Fanuc KAREL source: kt00881.KL

-- PROVISIONAL review KL for V770-1; original PC SHA256 7bfcebda0242e58e16e4d91c53400874c8d9c3006e6fad8e13b8db4fe4a92cd5
-- Incomplete behavior may be omitted. Consult companion uncertainty JSON. Do not deploy.
PROGRAM KT00881
%NOLOCKGROUP
VAR
  I1 : INTEGER
  I2 : INTEGER
  OUT : REAL
BEGIN
  -- UNRESOLVED_PC offsets 5-16; opcodes 2E,23
  -- UNRESOLVED_PC offsets 21-32; opcodes 2E,23
  -- UNRESOLVED_PC offsets 37-48; opcodes 2E,23
  -- UNRESOLVED_PC offsets 53-64; opcodes 2E,23
  -- UNRESOLVED_PC offsets 69-94; opcodes 27,27,21,64,27,21,64,76,23
  -- UNRESOLVED_PC offsets 99-103; opcodes 7F
END KT00881
